ABB RobotStudio station: Lab1.rsstnx

Station Lab1 (saved by RobotStudio 25.5.11605.0)
Controller IRB140_6_81
  mechanical unit ROB_1: IRB140_6_81_C_03, 6 joints, base frame (0, 0, 0) mm
Layout (positions relative to the parent item):
  - IRB140_6_81_C_03 [mechanism, from %ABB.RobotStudio.Models.IRB140%\IRB140_6_81_C_G_03.rslib] at (0, 0, 0) mm; joint values [0, 0, 0, 0, 0.5236, 0] (rad or m)
  - MyNewTool [mechanism] at (506.29, 0, 679.5) mm, rotated rx 180 ry 60 rz 180 deg
      TCP MyNewTool at (110.98, -0.23, 41.34) mm, rotated rx 0 ry -30 rz 180 deg
      links: Assembly 2
  - Pastel [part] at (327.56, -460.42, -59) mm, rotated rx 180 ry 0 rz -90 deg, size 150 x 200 x 50 mm
  - Banda [smart component]
      signals: DI DI_01, DI DI_02
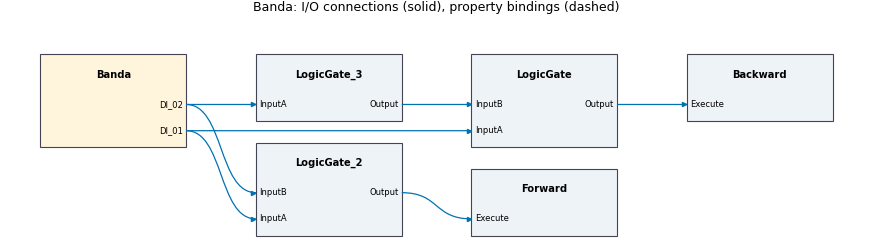
      connections:
        Banda.DI_02 -> LogicGate_3.InputA
        LogicGate_3.Output -> LogicGate.InputB
        LogicGate.Output -> Backward.Execute
        Banda.DI_02 -> LogicGate_2.InputB
        LogicGate_2.Output -> Forward.Execute
        Banda.DI_01 -> LogicGate_2.InputA
        Banda.DI_01 -> LogicGate.InputA
    - LogicGate [smart component, from Components\LogicGate.rslib]
        properties: Operator=AND; Delay=0.4
    - LogicGate_2 [smart component, from Components\LogicGate.rslib]
        properties: Operator=AND; Delay=0.4
    - LogicGate_3 [smart component, from Components\LogicGate.rslib]
        properties: Operator=NOT; Delay=0
    - Forward [smart component, from Components\LinearMover.rslib]
        properties: Object=Pastel; Direction=[0 -0.001 0]; Speed=0.328; Reference=Local; ReferenceObject=(none)
    - Backward [smart component, from Components\LinearMover.rslib]
        properties: Object=Pastel; Direction=[0 0.001 0]; Speed=0.328; Reference=Local; ReferenceObject=(none)
    - Start [smart component, from Components\Positioner.rslib] at (0, 0, 0) mm
        properties: Object=Pastel; Position=[-0.845372 -0.460416 -0.059]; Orientation=[3.14159265358979 0 -1.5707963267949]; Reference=Global; ReferenceObject=(none)
    - End [smart component, from Components\Positioner.rslib]
        properties: Object=Pastel; Position=[0.014628 -0.460416 -0.059]; Orientation=[3.14159265358979 0 -1.5707963267949]; Reference=Global; ReferenceObject=(none)
Attachment: MyNewTool is attached to IRB140_6_81_C_03 / Link6
Attachment: Start is attached to IRB140_6_81_C_03 / Link6
Station signals: DI DI_01, DI DI_02, DI DI_03
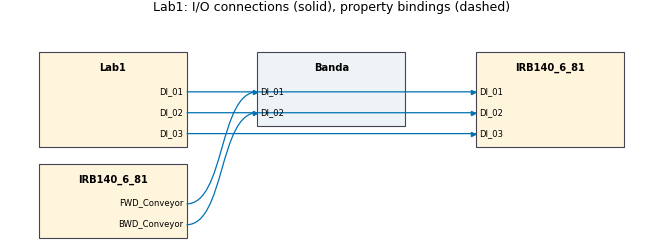
Station logic (signal -> signal, property => property):
  Lab1.DI_01 -> IRB140_6_81.DI_01
  Lab1.DI_02 -> IRB140_6_81.DI_02
  Lab1.DI_03 -> IRB140_6_81.DI_03
  IRB140_6_81.FWD_Conveyor -> Banda.DI_01
  IRB140_6_81.BWD_Conveyor -> Banda.DI_02
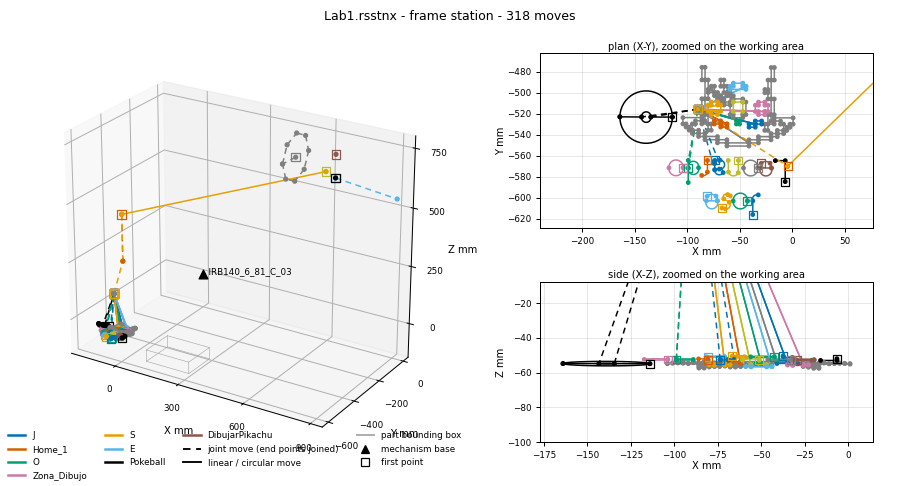
[picture p0: tool path of Lab1.rsstnx in frame station, 318 of 318 moves have a stored position in this frame; points joined in program order, loops and branches not executed]
Targets, tools, work objects and paths stored in the station, written as RAPID:
! task T_ROB1
MODULE Module1
  CONST robtarget E6_21:=[[119.525,55.911,0],[0,0,0,1],[0,0,0,0],[9E+09,9E+09,9E+09,9E+09,9E+09,9E+09]];
  PERS tooldata MyNewTool:=[TRUE,[[41.338,0.233,110.975],[0.866025404,0,0.5,0]],[1,[0,0,1],[1,0,0,0],0,0,0]];
  TASK PERS wobjdata Workobject_1:=[FALSE,TRUE,"",[[10.169850696,-448.889900169,-59],[0.018985691,0.705924683,-0.707820682,0.017313792]],[[0,0,0],[1,0,0,0]]];
  CONST robtarget D1:=[[123.545,108.722,0],[0,0,0,1],[-1,0,-1,1],[9E+09,9E+09,9E+09,9E+09,9E+09,9E+09]];
  CONST robtarget D2:=[[129.593,104.085,0],[0,0,0,1],[-1,0,-1,1],[9E+09,9E+09,9E+09,9E+09,9E+09,9E+09]];
  CONST robtarget D3:=[[123.185,98.948,0],[0,0,0,1],[-1,0,-1,1],[9E+09,9E+09,9E+09,9E+09,9E+09,9E+09]];
  CONST robtarget D4:=[[117.051,103.638,0],[0,0,0,1],[-1,0,-1,1],[9E+09,9E+09,9E+09,9E+09,9E+09,9E+09]];
  CONST robtarget Dibujo:=[[75,100,-150],[0,0,0,1],[-1,0,-1,1],[9E+09,9E+09,9E+09,9E+09,9E+09,9E+09]];
  CONST robtarget D5:=[[116.175,108.722,0],[0,0,0,1],[-1,0,-1,1],[9E+09,9E+09,9E+09,9E+09,9E+09,9E+09]];
  CONST robtarget D6:=[[137.325,108.722,0],[0,0,0,1],[-1,0,-1,1],[9E+09,9E+09,9E+09,9E+09,9E+09,9E+09]];
  CONST robtarget O1_2:=[[123.237,42.561,0],[0,0,0,1],[-1,0,-1,1],[9E+09,9E+09,9E+09,9E+09,9E+09,9E+09]];
  CONST robtarget O2_2:=[[130.813,49.503,0],[0,0,0,1],[-1,0,-1,1],[9E+09,9E+09,9E+09,9E+09,9E+09,9E+09]];
  CONST robtarget O3_2:=[[123.305,56.117,0],[0,0,0,1],[-1,0,-1,1],[9E+09,9E+09,9E+09,9E+09,9E+09,9E+09]];
  CONST robtarget O4_2:=[[115.831,49.349,0],[0,0,0,1],[-1,0,-1,1],[9E+09,9E+09,9E+09,9E+09,9E+09,9E+09]];
  CONST robtarget DibujoPk:=[[75,100,-150],[0,0,0,1],[0,0,0,0],[9E+09,9E+09,9E+09,9E+09,9E+09,9E+09]];
  CONST robtarget P2_1:=[[60.375,65.975,0],[0,0,0,1],[0,0,0,0],[9E+09,9E+09,9E+09,9E+09,9E+09,9E+09]];
  CONST robtarget P2_2:=[[60.375,56.975,0],[0,0,0,1],[0,0,0,0],[9E+09,9E+09,9E+09,9E+09,9E+09,9E+09]];
  CONST robtarget P2_3:=[[69.375,56.975,0],[0,0,0,1],[0,0,0,0],[9E+09,9E+09,9E+09,9E+09,9E+09,9E+09]];
  CONST robtarget P2_4:=[[69.375,65.975,0],[0,0,0,1],[0,0,0,0],[9E+09,9E+09,9E+09,9E+09,9E+09,9E+09]];
  CONST robtarget N1:=[[116.175,60.996,0],[0,0,0,1],[-1,0,-1,1],[9E+09,9E+09,9E+09,9E+09,9E+09,9E+09]];
  CONST robtarget N2:=[[127.893,61.049,0],[0,0,0,1],[-1,0,-1,1],[9E+09,9E+09,9E+09,9E+09,9E+09,9E+09]];
  CONST robtarget N3:=[[130.813,65.927,0],[0,0,0,1],[-1,0,-1,1],[9E+09,9E+09,9E+09,9E+09,9E+09,9E+09]];
  CONST robtarget N4:=[[127.169,70.439,0],[0,0,0,1],[-1,0,-1,1],[9E+09,9E+09,9E+09,9E+09,9E+09,9E+09]];
  CONST robtarget N5:=[[116.175,70.686,0],[0,0,0,1],[-1,0,-1,1],[9E+09,9E+09,9E+09,9E+09,9E+09,9E+09]];
  CONST robtarget P4_1:=[[81.375,71.975,0],[0,0,0,1],[0,0,0,0],[9E+09,9E+09,9E+09,9E+09,9E+09,9E+09]];
  CONST robtarget P4_2:=[[81.375,77.975,0],[0,0,0,1],[0,0,0,0],[9E+09,9E+09,9E+09,9E+09,9E+09,9E+09]];
  CONST robtarget P4_3:=[[78.375,77.975,0],[0,0,0,1],[0,0,0,0],[9E+09,9E+09,9E+09,9E+09,9E+09,9E+09]];
  CONST robtarget P4_4:=[[78.375,83.975,0],[0,0,0,1],[0,0,0,0],[9E+09,9E+09,9E+09,9E+09,9E+09,9E+09]];
  CONST robtarget P4_5:=[[81.375,83.975,0],[0,0,0,1],[0,0,0,0],[9E+09,9E+09,9E+09,9E+09,9E+09,9E+09]];
  CONST robtarget P4_6:=[[81.375,77.975,0],[0,0,0,1],[0,0,0,0],[9E+09,9E+09,9E+09,9E+09,9E+09,9E+09]];
  CONST robtarget P4_7:=[[84.375,77.975,0],[0,0,0,1],[0,0,0,0],[9E+09,9E+09,9E+09,9E+09,9E+09,9E+09]];
  CONST robtarget P4_8:=[[84.375,71.975,0],[0,0,0,1],[0,0,0,0],[9E+09,9E+09,9E+09,9E+09,9E+09,9E+09]];
  CONST robtarget P6_1:=[[69.375,35.975,0],[0,0,0,1],[0,0,0,0],[9E+09,9E+09,9E+09,9E+09,9E+09,9E+09]];
  CONST robtarget P6_2:=[[69.375,32.975,0],[0,0,0,1],[0,0,0,0],[9E+09,9E+09,9E+09,9E+09,9E+09,9E+09]];
  CONST robtarget P6_3:=[[63.375,32.975,0],[0,0,0,1],[0,0,0,0],[9E+09,9E+09,9E+09,9E+09,9E+09,9E+09]];
  CONST robtarget P6_4:=[[63.375,35.975,0],[0,0,0,1],[0,0,0,0],[9E+09,9E+09,9E+09,9E+09,9E+09,9E+09]];
  CONST robtarget P6_5:=[[60.375,35.975,0],[0,0,0,1],[0,0,0,0],[9E+09,9E+09,9E+09,9E+09,9E+09,9E+09]];
  CONST robtarget P6_6:=[[60.375,41.975,0],[0,0,0,1],[0,0,0,0],[9E+09,9E+09,9E+09,9E+09,9E+09,9E+09]];
  CONST robtarget P6_7:=[[63.375,41.975,0],[0,0,0,1],[0,0,0,0],[9E+09,9E+09,9E+09,9E+09,9E+09,9E+09]];
  CONST robtarget P6_8:=[[63.375,44.975,0],[0,0,0,1],[0,0,0,0],[9E+09,9E+09,9E+09,9E+09,9E+09,9E+09]];
  CONST robtarget P6_9:=[[69.375,44.975,0],[0,0,0,1],[0,0,0,0],[9E+09,9E+09,9E+09,9E+09,9E+09,9E+09]];
  CONST robtarget P6_10:=[[69.375,41.975,0],[0,0,0,1],[0,0,0,0],[9E+09,9E+09,9E+09,9E+09,9E+09,9E+09]];
  CONST robtarget P6_11:=[[72.375,41.975,0],[0,0,0,1],[0,0,0,0],[9E+09,9E+09,9E+09,9E+09,9E+09,9E+09]];
  CONST robtarget P6_12:=[[72.375,35.975,0],[0,0,0,1],[0,0,0,0],[9E+09,9E+09,9E+09,9E+09,9E+09,9E+09]];
  CONST robtarget O1_3:=[[123.237,113.603,0],[0,0,0,1],[-1,0,-1,1],[9E+09,9E+09,9E+09,9E+09,9E+09,9E+09]];
  CONST robtarget O2_3:=[[130.813,120.543,0],[0,0,0,1],[-1,0,-1,1],[9E+09,9E+09,9E+09,9E+09,9E+09,9E+09]];
  CONST robtarget O3_3:=[[123.305,127.159,0],[0,0,0,1],[-1,0,-1,1],[9E+09,9E+09,9E+09,9E+09,9E+09,9E+09]];
  CONST robtarget O4_3:=[[115.831,120.388,0],[0,0,0,1],[-1,0,-1,1],[9E+09,9E+09,9E+09,9E+09,9E+09,9E+09]];
  CONST robtarget PB1:=[[74.913,124.015,0],[0,0,0,1],[-1,0,-1,1],[9E+09,9E+09,9E+09,9E+09,9E+09,9E+09]];
  CONST robtarget PB2:=[[100,149.015,0],[0,0,0,1],[-1,0,-1,1],[9E+09,9E+09,9E+09,9E+09,9E+09,9E+09]];
  CONST robtarget PB3:=[[74.812,174.015,0],[0,0,0,1],[-1,0,-1,1],[9E+09,9E+09,9E+09,9E+09,9E+09,9E+09]];
  CONST robtarget PB4:=[[50,149.015,0],[0,0,0,1],[-1,0,-1,1],[9E+09,9E+09,9E+09,9E+09,9E+09,9E+09]];
  CONST robtarget PB5:=[[74.913,144.515,0],[0,0,0,1],[-1,0,-1,1],[9E+09,9E+09,9E+09,9E+09,9E+09,9E+09]];
  CONST robtarget PB6:=[[80,149.015,0],[0,0,0,1],[-1,0,-1,1],[9E+09,9E+09,9E+09,9E+09,9E+09,9E+09]];
  CONST robtarget PB7:=[[74.913,153.345,0],[0,0,0,1],[-1,0,-1,1],[9E+09,9E+09,9E+09,9E+09,9E+09,9E+09]];
  CONST robtarget PB8:=[[70,149.015,0],[0,0,0,1],[-1,0,-1,1],[9E+09,9E+09,9E+09,9E+09,9E+09,9E+09]];
  CONST robtarget J1:=[[167.685,47.174,0],[0,0,0,1],[-1,0,-1,1],[9E+09,9E+09,9E+09,9E+09,9E+09,9E+09]];
  CONST robtarget J2:=[[154.611,47.174,0],[0,0,0,1],[-1,0,-1,1],[9E+09,9E+09,9E+09,9E+09,9E+09,9E+09]];
  CONST robtarget J3:=[[150.083,46.324,0],[0,0,0,1],[-1,0,-1,1],[9E+09,9E+09,9E+09,9E+09,9E+09,9E+09]];
  CONST robtarget J4:=[[148.923,41.986,0],[0,0,0,1],[-1,0,-1,1],[9E+09,9E+09,9E+09,9E+09,9E+09,9E+09]];
  CONST robtarget P8_1:=[[45.375,53.975,0],[0,0,0,1],[0,0,0,0],[9E+09,9E+09,9E+09,9E+09,9E+09,9E+09]];
  CONST robtarget P8_2:=[[45.375,56.975,0],[0,0,0,1],[0,0,0,0],[9E+09,9E+09,9E+09,9E+09,9E+09,9E+09]];
  CONST robtarget P8_3:=[[42.375,56.975,0],[0,0,0,1],[0,0,0,0],[9E+09,9E+09,9E+09,9E+09,9E+09,9E+09]];
  CONST robtarget P8_4:=[[42.375,65.975,0],[0,0,0,1],[0,0,0,0],[9E+09,9E+09,9E+09,9E+09,9E+09,9E+09]];
  CONST robtarget P8_5:=[[45.375,65.975,0],[0,0,0,1],[0,0,0,0],[9E+09,9E+09,9E+09,9E+09,9E+09,9E+09]];
  CONST robtarget P8_6:=[[45.375,68.975,0],[0,0,0,1],[0,0,0,0],[9E+09,9E+09,9E+09,9E+09,9E+09,9E+09]];
  CONST robtarget P8_7:=[[48.375,68.975,0],[0,0,0,1],[0,0,0,0],[9E+09,9E+09,9E+09,9E+09,9E+09,9E+09]];
  CONST robtarget P8_8:=[[48.375,53.975,0],[0,0,0,1],[0,0,0,0],[9E+09,9E+09,9E+09,9E+09,9E+09,9E+09]];
  CONST robtarget wobjreal:=[[10.17,-448.89,43.77],[0.275144,0.645288,0.659942,-0.269026],[-1,0,0,1],[9E+09,9E+09,9E+09,9E+09,9E+09,9E+09]];
  CONST robtarget P1_1:=[[99.375,50.975,0],[0,0,0,1],[0,0,0,0],[9E+09,9E+09,9E+09,9E+09,9E+09,9E+09]];
  CONST robtarget P1_2:=[[99.375,41.975,0],[0,0,0,1],[0,0,0,0],[9E+09,9E+09,9E+09,9E+09,9E+09,9E+09]];
  CONST robtarget P1_3:=[[96.375,41.975,0],[0,0,0,1],[0,0,0,0],[9E+09,9E+09,9E+09,9E+09,9E+09,9E+09]];
  CONST robtarget P1_4:=[[96.375,29.975,0],[0,0,0,1],[0,0,0,0],[9E+09,9E+09,9E+09,9E+09,9E+09,9E+09]];
  CONST robtarget P1_5:=[[93.375,29.975,0],[0,0,0,1],[0,0,0,0],[9E+09,9E+09,9E+09,9E+09,9E+09,9E+09]];
  CONST robtarget P1_6:=[[93.375,23.975,0],[0,0,0,1],[0,0,0,0],[9E+09,9E+09,9E+09,9E+09,9E+09,9E+09]];
  CONST robtarget P1_7:=[[90.375,23.975,0],[0,0,0,1],[0,0,0,0],[9E+09,9E+09,9E+09,9E+09,9E+09,9E+09]];
  CONST robtarget P1_8:=[[90.375,17.975,0],[0,0,0,1],[0,0,0,0],[9E+09,9E+09,9E+09,9E+09,9E+09,9E+09]];
  CONST robtarget P1_9:=[[87.375,17.975,0],[0,0,0,1],[0,0,0,0],[9E+09,9E+09,9E+09,9E+09,9E+09,9E+09]];
  CONST robtarget P1_10:=[[87.375,14.975,0],[0,0,0,1],[0,0,0,0],[9E+09,9E+09,9E+09,9E+09,9E+09,9E+09]];
  CONST robtarget P1_11:=[[84.375,14.975,0],[0,0,0,1],[0,0,0,0],[9E+09,9E+09,9E+09,9E+09,9E+09,9E+09]];
  CONST robtarget P1_12:=[[84.375,11.975,0],[0,0,0,1],[0,0,0,0],[9E+09,9E+09,9E+09,9E+09,9E+09,9E+09]];
  CONST robtarget P1_13:=[[81.375,11.975,0],[0,0,0,1],[0,0,0,0],[9E+09,9E+09,9E+09,9E+09,9E+09,9E+09]];
  CONST robtarget P1_14:=[[81.375,8.975,0],[0,0,0,1],[0,0,0,0],[9E+09,9E+09,9E+09,9E+09,9E+09,9E+09]];
  CONST robtarget P1_15:=[[75.375,8.975,0],[0,0,0,1],[0,0,0,0],[9E+09,9E+09,9E+09,9E+09,9E+09,9E+09]];
  CONST robtarget P1_16:=[[75.375,26.975,0],[0,0,0,1],[0,0,0,0],[9E+09,9E+09,9E+09,9E+09,9E+09,9E+09]];
  CONST robtarget P1_17:=[[78.375,26.975,0],[0,0,0,1],[0,0,0,0],[9E+09,9E+09,9E+09,9E+09,9E+09,9E+09]];
  CONST robtarget P1_18:=[[78.375,29.975,0],[0,0,0,1],[0,0,0,0],[9E+09,9E+09,9E+09,9E+09,9E+09,9E+09]];
  CONST robtarget P1_19:=[[72.375,29.975,0],[0,0,0,1],[0,0,0,0],[9E+09,9E+09,9E+09,9E+09,9E+09,9E+09]];
  CONST robtarget P1_20:=[[72.375,26.975,0],[0,0,0,1],[0,0,0,0],[9E+09,9E+09,9E+09,9E+09,9E+09,9E+09]];
  CONST robtarget P1_21:=[[57.375,26.975,0],[0,0,0,1],[0,0,0,0],[9E+09,9E+09,9E+09,9E+09,9E+09,9E+09]];
  CONST robtarget P1_22:=[[57.375,29.975,0],[0,0,0,1],[0,0,0,0],[9E+09,9E+09,9E+09,9E+09,9E+09,9E+09]];
  CONST robtarget P1_23:=[[39.375,29.975,0],[0,0,0,1],[0,0,0,0],[9E+09,9E+09,9E+09,9E+09,9E+09,9E+09]];
  CONST robtarget P1_24:=[[39.375,26.975,0],[0,0,0,1],[0,0,0,0],[9E+09,9E+09,9E+09,9E+09,9E+09,9E+09]];
  CONST robtarget P1_25:=[[27.375,26.975,0],[0,0,0,1],[0,0,0,0],[9E+09,9E+09,9E+09,9E+09,9E+09,9E+09]];
  CONST robtarget P1_26:=[[27.375,29.975,0],[0,0,0,1],[0,0,0,0],[9E+09,9E+09,9E+09,9E+09,9E+09,9E+09]];
  CONST robtarget P1_27:=[[39.375,29.975,0],[0,0,0,1],[0,0,0,0],[9E+09,9E+09,9E+09,9E+09,9E+09,9E+09]];
  CONST robtarget P1_28:=[[39.375,32.975,0],[0,0,0,1],[0,0,0,0],[9E+09,9E+09,9E+09,9E+09,9E+09,9E+09]];
  CONST robtarget P1_29:=[[48.375,32.975,0],[0,0,0,1],[0,0,0,0],[9E+09,9E+09,9E+09,9E+09,9E+09,9E+09]];
  CONST robtarget P1_30:=[[48.375,35.975,0],[0,0,0,1],[0,0,0,0],[9E+09,9E+09,9E+09,9E+09,9E+09,9E+09]];
  CONST robtarget P1_31:=[[51.375,35.975,0],[0,0,0,1],[0,0,0,0],[9E+09,9E+09,9E+09,9E+09,9E+09,9E+09]];
  CONST robtarget P1_32:=[[51.375,32.975,0],[0,0,0,1],[0,0,0,0],[9E+09,9E+09,9E+09,9E+09,9E+09,9E+09]];
  CONST robtarget P1_33:=[[57.375,32.975,0],[0,0,0,1],[0,0,0,0],[9E+09,9E+09,9E+09,9E+09,9E+09,9E+09]];
  CONST robtarget P1_34:=[[57.375,29.975,0],[0,0,0,1],[0,0,0,0],[9E+09,9E+09,9E+09,9E+09,9E+09,9E+09]];
  CONST robtarget P1_35:=[[72.375,29.975,0],[0,0,0,1],[0,0,0,0],[9E+09,9E+09,9E+09,9E+09,9E+09,9E+09]];
  CONST robtarget P1_36:=[[72.375,32.975,0],[0,0,0,1],[0,0,0,0],[9E+09,9E+09,9E+09,9E+09,9E+09,9E+09]];
  CONST robtarget P1_37:=[[81.375,32.975,0],[0,0,0,1],[0,0,0,0],[9E+09,9E+09,9E+09,9E+09,9E+09,9E+09]];
  CONST robtarget P1_38:=[[81.375,35.975,0],[0,0,0,1],[0,0,0,0],[9E+09,9E+09,9E+09,9E+09,9E+09,9E+09]];
  CONST robtarget P1_39:=[[87.375,35.975,0],[0,0,0,1],[0,0,0,0],[9E+09,9E+09,9E+09,9E+09,9E+09,9E+09]];
  CONST robtarget P1_40:=[[87.375,32.975,0],[0,0,0,1],[0,0,0,0],[9E+09,9E+09,9E+09,9E+09,9E+09,9E+09]];
  CONST robtarget P1_41:=[[81.375,32.975,0],[0,0,0,1],[0,0,0,0],[9E+09,9E+09,9E+09,9E+09,9E+09,9E+09]];
  CONST robtarget P1_42:=[[81.375,26.975,0],[0,0,0,1],[0,0,0,0],[9E+09,9E+09,9E+09,9E+09,9E+09,9E+09]];
  CONST robtarget P1_43:=[[78.375,26.975,0],[0,0,0,1],[0,0,0,0],[9E+09,9E+09,9E+09,9E+09,9E+09,9E+09]];
  CONST robtarget P1_44:=[[78.375,20.975,0],[0,0,0,1],[0,0,0,0],[9E+09,9E+09,9E+09,9E+09,9E+09,9E+09]];
  CONST robtarget P1_45:=[[81.375,20.975,0],[0,0,0,1],[0,0,0,0],[9E+09,9E+09,9E+09,9E+09,9E+09,9E+09]];
  CONST robtarget P1_46:=[[81.375,17.975,0],[0,0,0,1],[0,0,0,0],[9E+09,9E+09,9E+09,9E+09,9E+09,9E+09]];
  CONST robtarget P1_47:=[[87.375,17.975,0],[0,0,0,1],[0,0,0,0],[9E+09,9E+09,9E+09,9E+09,9E+09,9E+09]];
  CONST robtarget P1_48:=[[87.375,23.975,0],[0,0,0,1],[0,0,0,0],[9E+09,9E+09,9E+09,9E+09,9E+09,9E+09]];
  CONST robtarget P1_49:=[[90.375,23.975,0],[0,0,0,1],[0,0,0,0],[9E+09,9E+09,9E+09,9E+09,9E+09,9E+09]];
  CONST robtarget P1_50:=[[90.375,29.975,0],[0,0,0,1],[0,0,0,0],[9E+09,9E+09,9E+09,9E+09,9E+09,9E+09]];
  CONST robtarget P1_51:=[[93.375,29.975,0],[0,0,0,1],[0,0,0,0],[9E+09,9E+09,9E+09,9E+09,9E+09,9E+09]];
  CONST robtarget P1_52:=[[93.375,41.975,0],[0,0,0,1],[0,0,0,0],[9E+09,9E+09,9E+09,9E+09,9E+09,9E+09]];
  CONST robtarget P1_53:=[[96.375,41.975,0],[0,0,0,1],[0,0,0,0],[9E+09,9E+09,9E+09,9E+09,9E+09,9E+09]];
  CONST robtarget P1_54:=[[96.375,50.975,0],[0,0,0,1],[0,0,0,0],[9E+09,9E+09,9E+09,9E+09,9E+09,9E+09]];
  CONST robtarget P1_55:=[[99.375,50.975,0],[0,0,0,1],[0,0,0,0],[9E+09,9E+09,9E+09,9E+09,9E+09,9E+09]];
  CONST robtarget P1_56:=[[99.375,71.975,0],[0,0,0,1],[0,0,0,0],[9E+09,9E+09,9E+09,9E+09,9E+09,9E+09]];
  CONST robtarget P1_57:=[[96.375,71.975,0],[0,0,0,1],[0,0,0,0],[9E+09,9E+09,9E+09,9E+09,9E+09,9E+09]];
  CONST robtarget P1_58:=[[96.375,80.975,0],[0,0,0,1],[0,0,0,0],[9E+09,9E+09,9E+09,9E+09,9E+09,9E+09]];
  CONST robtarget P1_59:=[[93.375,80.975,0],[0,0,0,1],[0,0,0,0],[9E+09,9E+09,9E+09,9E+09,9E+09,9E+09]];
  CONST robtarget P1_60:=[[93.375,92.975,0],[0,0,0,1],[0,0,0,0],[9E+09,9E+09,9E+09,9E+09,9E+09,9E+09]];
  CONST robtarget P1_61:=[[90.375,92.975,0],[0,0,0,1],[0,0,0,0],[9E+09,9E+09,9E+09,9E+09,9E+09,9E+09]];
  CONST robtarget P1_62:=[[90.375,98.975,0],[0,0,0,1],[0,0,0,0],[9E+09,9E+09,9E+09,9E+09,9E+09,9E+09]];
  CONST robtarget P1_63:=[[87.375,98.975,0],[0,0,0,1],[0,0,0,0],[9E+09,9E+09,9E+09,9E+09,9E+09,9E+09]];
  CONST robtarget P1_64:=[[87.375,104.975,0],[0,0,0,1],[0,0,0,0],[9E+09,9E+09,9E+09,9E+09,9E+09,9E+09]];
  CONST robtarget P1_65:=[[81.375,104.975,0],[0,0,0,1],[0,0,0,0],[9E+09,9E+09,9E+09,9E+09,9E+09,9E+09]];
  CONST robtarget P1_66:=[[81.375,101.975,0],[0,0,0,1],[0,0,0,0],[9E+09,9E+09,9E+09,9E+09,9E+09,9E+09]];
  CONST robtarget P1_67:=[[78.375,101.975,0],[0,0,0,1],[0,0,0,0],[9E+09,9E+09,9E+09,9E+09,9E+09,9E+09]];
  CONST robtarget P1_68:=[[78.375,95.975,0],[0,0,0,1],[0,0,0,0],[9E+09,9E+09,9E+09,9E+09,9E+09,9E+09]];
  CONST robtarget P1_69:=[[81.375,95.975,0],[0,0,0,1],[0,0,0,0],[9E+09,9E+09,9E+09,9E+09,9E+09,9E+09]];
  CONST robtarget P1_70:=[[81.375,89.975,0],[0,0,0,1],[0,0,0,0],[9E+09,9E+09,9E+09,9E+09,9E+09,9E+09]];
  CONST robtarget P1_71:=[[87.375,89.975,0],[0,0,0,1],[0,0,0,0],[9E+09,9E+09,9E+09,9E+09,9E+09,9E+09]];
  CONST robtarget P1_72:=[[87.375,86.975,0],[0,0,0,1],[0,0,0,0],[9E+09,9E+09,9E+09,9E+09,9E+09,9E+09]];
  CONST robtarget P1_73:=[[81.375,86.975,0],[0,0,0,1],[0,0,0,0],[9E+09,9E+09,9E+09,9E+09,9E+09,9E+09]];
  CONST robtarget P1_74:=[[81.375,89.975,0],[0,0,0,1],[0,0,0,0],[9E+09,9E+09,9E+09,9E+09,9E+09,9E+09]];
  CONST robtarget P1_75:=[[72.375,89.975,0],[0,0,0,1],[0,0,0,0],[9E+09,9E+09,9E+09,9E+09,9E+09,9E+09]];
  CONST robtarget P1_76:=[[72.375,92.975,0],[0,0,0,1],[0,0,0,0],[9E+09,9E+09,9E+09,9E+09,9E+09,9E+09]];
  CONST robtarget P1_77:=[[57.375,92.975,0],[0,0,0,1],[0,0,0,0],[9E+09,9E+09,9E+09,9E+09,9E+09,9E+09]];
  CONST robtarget P1_78:=[[57.375,89.975,0],[0,0,0,1],[0,0,0,0],[9E+09,9E+09,9E+09,9E+09,9E+09,9E+09]];
  CONST robtarget P1_79:=[[51.375,89.975,0],[0,0,0,1],[0,0,0,0],[9E+09,9E+09,9E+09,9E+09,9E+09,9E+09]];
  CONST robtarget P1_80:=[[51.375,83.975,0],[0,0,0,1],[0,0,0,0],[9E+09,9E+09,9E+09,9E+09,9E+09,9E+09]];
  CONST robtarget P1_81:=[[54.375,83.975,0],[0,0,0,1],[0,0,0,0],[9E+09,9E+09,9E+09,9E+09,9E+09,9E+09]];
  CONST robtarget P1_82:=[[54.375,80.975,0],[0,0,0,1],[0,0,0,0],[9E+09,9E+09,9E+09,9E+09,9E+09,9E+09]];
  CONST robtarget P1_83:=[[57.375,80.975,0],[0,0,0,1],[0,0,0,0],[9E+09,9E+09,9E+09,9E+09,9E+09,9E+09]];
  CONST robtarget P1_84:=[[57.375,77.975,0],[0,0,0,1],[0,0,0,0],[9E+09,9E+09,9E+09,9E+09,9E+09,9E+09]];
  CONST robtarget P1_85:=[[60.375,77.975,0],[0,0,0,1],[0,0,0,0],[9E+09,9E+09,9E+09,9E+09,9E+09,9E+09]];
  CONST robtarget P1_86:=[[60.375,74.975,0],[0,0,0,1],[0,0,0,0],[9E+09,9E+09,9E+09,9E+09,9E+09,9E+09]];
  CONST robtarget P1_87:=[[63.375,74.975,0],[0,0,0,1],[0,0,0,0],[9E+09,9E+09,9E+09,9E+09,9E+09,9E+09]];
  CONST robtarget P1_88:=[[63.375,68.975,0],[0,0,0,1],[0,0,0,0],[9E+09,9E+09,9E+09,9E+09,9E+09,9E+09]];
  CONST robtarget P1_89:=[[72.375,68.975,0],[0,0,0,1],[0,0,0,0],[9E+09,9E+09,9E+09,9E+09,9E+09,9E+09]];
  CONST robtarget P1_90:=[[72.375,65.975,0],[0,0,0,1],[0,0,0,0],[9E+09,9E+09,9E+09,9E+09,9E+09,9E+09]];
  CONST robtarget P1_91:=[[75.375,65.975,0],[0,0,0,1],[0,0,0,0],[9E+09,9E+09,9E+09,9E+09,9E+09,9E+09]];
  CONST robtarget P1_92:=[[75.375,56.975,0],[0,0,0,1],[0,0,0,0],[9E+09,9E+09,9E+09,9E+09,9E+09,9E+09]];
  CONST robtarget P1_93:=[[72.375,56.975,0],[0,0,0,1],[0,0,0,0],[9E+09,9E+09,9E+09,9E+09,9E+09,9E+09]];
  CONST robtarget P1_94:=[[72.375,53.975,0],[0,0,0,1],[0,0,0,0],[9E+09,9E+09,9E+09,9E+09,9E+09,9E+09]];
  CONST robtarget P1_95:=[[60.375,53.975,0],[0,0,0,1],[0,0,0,0],[9E+09,9E+09,9E+09,9E+09,9E+09,9E+09]];
  CONST robtarget P1_96:=[[60.375,56.975,0],[0,0,0,1],[0,0,0,0],[9E+09,9E+09,9E+09,9E+09,9E+09,9E+09]];
  CONST robtarget P1_97:=[[57.375,56.975,0],[0,0,0,1],[0,0,0,0],[9E+09,9E+09,9E+09,9E+09,9E+09,9E+09]];
  CONST robtarget P1_98:=[[57.375,65.975,0],[0,0,0,1],[0,0,0,0],[9E+09,9E+09,9E+09,9E+09,9E+09,9E+09]];
  CONST robtarget P1_99:=[[54.375,65.975,0],[0,0,0,1],[0,0,0,0],[9E+09,9E+09,9E+09,9E+09,9E+09,9E+09]];
  CONST robtarget P1_100:=[[54.375,68.975,0],[0,0,0,1],[0,0,0,0],[9E+09,9E+09,9E+09,9E+09,9E+09,9E+09]];
  CONST robtarget P1_101:=[[51.375,68.975,0],[0,0,0,1],[0,0,0,0],[9E+09,9E+09,9E+09,9E+09,9E+09,9E+09]];
  CONST robtarget P1_102:=[[51.375,71.975,0],[0,0,0,1],[0,0,0,0],[9E+09,9E+09,9E+09,9E+09,9E+09,9E+09]];
  CONST robtarget P1_103:=[[45.375,71.975,0],[0,0,0,1],[0,0,0,0],[9E+09,9E+09,9E+09,9E+09,9E+09,9E+09]];
  CONST robtarget P1_104:=[[45.375,74.975,0],[0,0,0,1],[0,0,0,0],[9E+09,9E+09,9E+09,9E+09,9E+09,9E+09]];
  CONST robtarget P1_105:=[[39.375,74.975,0],[0,0,0,1],[0,0,0,0],[9E+09,9E+09,9E+09,9E+09,9E+09,9E+09]];
  CONST robtarget P1_106:=[[39.375,77.975,0],[0,0,0,1],[0,0,0,0],[9E+09,9E+09,9E+09,9E+09,9E+09,9E+09]];
  CONST robtarget P1_107:=[[45.375,77.975,0],[0,0,0,1],[0,0,0,0],[9E+09,9E+09,9E+09,9E+09,9E+09,9E+09]];
  CONST robtarget P1_108:=[[45.375,74.975,0],[0,0,0,1],[0,0,0,0],[9E+09,9E+09,9E+09,9E+09,9E+09,9E+09]];
  CONST robtarget P1_109:=[[51.375,74.975,0],[0,0,0,1],[0,0,0,0],[9E+09,9E+09,9E+09,9E+09,9E+09,9E+09]];
  CONST robtarget P1_110:=[[51.375,71.975,0],[0,0,0,1],[0,0,0,0],[9E+09,9E+09,9E+09,9E+09,9E+09,9E+09]];
  CONST robtarget P1_111:=[[54.375,71.975,0],[0,0,0,1],[0,0,0,0],[9E+09,9E+09,9E+09,9E+09,9E+09,9E+09]];
  CONST robtarget P1_112:=[[54.375,68.975,0],[0,0,0,1],[0,0,0,0],[9E+09,9E+09,9E+09,9E+09,9E+09,9E+09]];
  CONST robtarget P1_113:=[[60.375,68.975,0],[0,0,0,1],[0,0,0,0],[9E+09,9E+09,9E+09,9E+09,9E+09,9E+09]];
  CONST robtarget P1_114:=[[60.375,74.975,0],[0,0,0,1],[0,0,0,0],[9E+09,9E+09,9E+09,9E+09,9E+09,9E+09]];
  CONST robtarget P1_115:=[[57.375,74.975,0],[0,0,0,1],[0,0,0,0],[9E+09,9E+09,9E+09,9E+09,9E+09,9E+09]];
  CONST robtarget P1_116:=[[57.375,77.975,0],[0,0,0,1],[0,0,0,0],[9E+09,9E+09,9E+09,9E+09,9E+09,9E+09]];
  CONST robtarget P1_117:=[[54.375,77.975,0],[0,0,0,1],[0,0,0,0],[9E+09,9E+09,9E+09,9E+09,9E+09,9E+09]];
  CONST robtarget P1_118:=[[54.375,80.975,0],[0,0,0,1],[0,0,0,0],[9E+09,9E+09,9E+09,9E+09,9E+09,9E+09]];
  CONST robtarget P1_119:=[[51.375,80.975,0],[0,0,0,1],[0,0,0,0],[9E+09,9E+09,9E+09,9E+09,9E+09,9E+09]];
  CONST robtarget P1_120:=[[51.375,83.975,0],[0,0,0,1],[0,0,0,0],[9E+09,9E+09,9E+09,9E+09,9E+09,9E+09]];
  CONST robtarget P1_121:=[[45.375,83.975,0],[0,0,0,1],[0,0,0,0],[9E+09,9E+09,9E+09,9E+09,9E+09,9E+09]];
  CONST robtarget P1_122:=[[45.375,86.975,0],[0,0,0,1],[0,0,0,0],[9E+09,9E+09,9E+09,9E+09,9E+09,9E+09]];
  CONST robtarget P1_123:=[[48.375,86.975,0],[0,0,0,1],[0,0,0,0],[9E+09,9E+09,9E+09,9E+09,9E+09,9E+09]];
  CONST robtarget P1_124:=[[48.375,89.975,0],[0,0,0,1],[0,0,0,0],[9E+09,9E+09,9E+09,9E+09,9E+09,9E+09]];
  CONST robtarget P1_125:=[[39.375,89.975,0],[0,0,0,1],[0,0,0,0],[9E+09,9E+09,9E+09,9E+09,9E+09,9E+09]];
  CONST robtarget P1_126:=[[39.375,92.975,0],[0,0,0,1],[0,0,0,0],[9E+09,9E+09,9E+09,9E+09,9E+09,9E+09]];
  CONST robtarget P1_127:=[[27.375,92.975,0],[0,0,0,1],[0,0,0,0],[9E+09,9E+09,9E+09,9E+09,9E+09,9E+09]];
  CONST robtarget P1_128:=[[27.375,95.975,0],[0,0,0,1],[0,0,0,0],[9E+09,9E+09,9E+09,9E+09,9E+09,9E+09]];
  CONST robtarget P1_129:=[[39.375,95.975,0],[0,0,0,1],[0,0,0,0],[9E+09,9E+09,9E+09,9E+09,9E+09,9E+09]];
  CONST robtarget P1_130:=[[39.375,92.975,0],[0,0,0,1],[0,0,0,0],[9E+09,9E+09,9E+09,9E+09,9E+09,9E+09]];
  CONST robtarget P1_131:=[[57.375,92.975,0],[0,0,0,1],[0,0,0,0],[9E+09,9E+09,9E+09,9E+09,9E+09,9E+09]];
  CONST robtarget P1_132:=[[57.375,95.975,0],[0,0,0,1],[0,0,0,0],[9E+09,9E+09,9E+09,9E+09,9E+09,9E+09]];
  CONST robtarget P1_133:=[[72.375,95.975,0],[0,0,0,1],[0,0,0,0],[9E+09,9E+09,9E+09,9E+09,9E+09,9E+09]];
  CONST robtarget P1_134:=[[72.375,92.975,0],[0,0,0,1],[0,0,0,0],[9E+09,9E+09,9E+09,9E+09,9E+09,9E+09]];
  CONST robtarget P1_135:=[[78.375,92.975,0],[0,0,0,1],[0,0,0,0],[9E+09,9E+09,9E+09,9E+09,9E+09,9E+09]];
  CONST robtarget P1_136:=[[78.375,95.975,0],[0,0,0,1],[0,0,0,0],[9E+09,9E+09,9E+09,9E+09,9E+09,9E+09]];
  CONST robtarget P1_137:=[[75.375,95.975,0],[0,0,0,1],[0,0,0,0],[9E+09,9E+09,9E+09,9E+09,9E+09,9E+09]];
  CONST robtarget P1_138:=[[75.375,113.975,0],[0,0,0,1],[0,0,0,0],[9E+09,9E+09,9E+09,9E+09,9E+09,9E+09]];
  CONST robtarget P1_139:=[[81.375,113.975,0],[0,0,0,1],[0,0,0,0],[9E+09,9E+09,9E+09,9E+09,9E+09,9E+09]];
  CONST robtarget P1_140:=[[81.375,110.975,0],[0,0,0,1],[0,0,0,0],[9E+09,9E+09,9E+09,9E+09,9E+09,9E+09]];
  CONST robtarget P1_141:=[[84.375,110.975,0],[0,0,0,1],[0,0,0,0],[9E+09,9E+09,9E+09,9E+09,9E+09,9E+09]];
  CONST robtarget P1_142:=[[84.375,107.975,0],[0,0,0,1],[0,0,0,0],[9E+09,9E+09,9E+09,9E+09,9E+09,9E+09]];
  CONST robtarget P1_143:=[[87.375,107.975,0],[0,0,0,1],[0,0,0,0],[9E+09,9E+09,9E+09,9E+09,9E+09,9E+09]];
  CONST robtarget P1_144:=[[87.375,104.975,0],[0,0,0,1],[0,0,0,0],[9E+09,9E+09,9E+09,9E+09,9E+09,9E+09]];
  CONST robtarget P1_145:=[[90.375,104.975,0],[0,0,0,1],[0,0,0,0],[9E+09,9E+09,9E+09,9E+09,9E+09,9E+09]];
  CONST robtarget P1_146:=[[90.375,98.975,0],[0,0,0,1],[0,0,0,0],[9E+09,9E+09,9E+09,9E+09,9E+09,9E+09]];
  CONST robtarget P1_147:=[[93.375,98.975,0],[0,0,0,1],[0,0,0,0],[9E+09,9E+09,9E+09,9E+09,9E+09,9E+09]];
  CONST robtarget P1_148:=[[93.375,92.975,0],[0,0,0,1],[0,0,0,0],[9E+09,9E+09,9E+09,9E+09,9E+09,9E+09]];
  CONST robtarget P1_149:=[[96.375,92.975,0],[0,0,0,1],[0,0,0,0],[9E+09,9E+09,9E+09,9E+09,9E+09,9E+09]];
  CONST robtarget P1_150:=[[96.375,80.975,0],[0,0,0,1],[0,0,0,0],[9E+09,9E+09,9E+09,9E+09,9E+09,9E+09]];
  CONST robtarget P1_151:=[[99.375,80.975,0],[0,0,0,1],[0,0,0,0],[9E+09,9E+09,9E+09,9E+09,9E+09,9E+09]];
  CONST robtarget P1_152:=[[99.375,71.975,0],[0,0,0,1],[0,0,0,0],[9E+09,9E+09,9E+09,9E+09,9E+09,9E+09]];
  CONST robtarget P1_153:=[[102.375,71.975,0],[0,0,0,1],[0,0,0,0],[9E+09,9E+09,9E+09,9E+09,9E+09,9E+09]];
  CONST robtarget P1_154:=[[102.375,50.975,0],[0,0,0,1],[0,0,0,0],[9E+09,9E+09,9E+09,9E+09,9E+09,9E+09]];
  CONST robtarget A1:=[[116.175,83.52,0],[0,0,0,1],[-1,0,-1,1],[9E+09,9E+09,9E+09,9E+09,9E+09,9E+09]];
  CONST robtarget A2:=[[125.057,83.52,0],[0,0,0,1],[-1,0,-1,1],[9E+09,9E+09,9E+09,9E+09,9E+09,9E+09]];
  CONST robtarget A3:=[[129.549,80.727,0],[0,0,0,1],[-1,0,-1,1],[9E+09,9E+09,9E+09,9E+09,9E+09,9E+09]];
  CONST robtarget A4:=[[127.721,75.478,0],[0,0,0,1],[-1,0,-1,1],[9E+09,9E+09,9E+09,9E+09,9E+09,9E+09]];
  CONST robtarget A5:=[[124.405,79.121,0],[0,0,0,1],[-1,0,-1,1],[9E+09,9E+09,9E+09,9E+09,9E+09,9E+09]];
  CONST robtarget A6:=[[119.869,74.173,0],[0,0,0,1],[-1,0,-1,1],[9E+09,9E+09,9E+09,9E+09,9E+09,9E+09]];
  CONST robtarget A7:=[[115.831,78.607,0],[0,0,0,1],[-1,0,-1,1],[9E+09,9E+09,9E+09,9E+09,9E+09,9E+09]];
  CONST robtarget A8:=[[116.673,81.448,0],[0,0,0,1],[-1,0,-1,1],[9E+09,9E+09,9E+09,9E+09,9E+09,9E+09]];
  CONST robtarget A9:=[[119.011,83.469,0],[0,0,0,1],[-1,0,-1,1],[9E+09,9E+09,9E+09,9E+09,9E+09,9E+09]];
  CONST robtarget L1:=[[136.191,16.345,0],[0,0,0,1],[-1,0,-1,1],[9E+09,9E+09,9E+09,9E+09,9E+09,9E+09]];
  CONST robtarget L2:=[[116.175,16.345,0],[0,0,0,1],[-1,0,-1,1],[9E+09,9E+09,9E+09,9E+09,9E+09,9E+09]];
  CONST robtarget L3:=[[116.175,25.793,0],[0,0,0,1],[-1,0,-1,1],[9E+09,9E+09,9E+09,9E+09,9E+09,9E+09]];
  CONST robtarget R1:=[[116.175,90.46,0],[0,0,0,1],[-1,0,-1,1],[9E+09,9E+09,9E+09,9E+09,9E+09,9E+09]];
  CONST robtarget R2:=[[127.309,90.513,0],[0,0,0,1],[-1,0,-1,1],[9E+09,9E+09,9E+09,9E+09,9E+09,9E+09]];
  CONST robtarget R2_2:=[[130.135,92.453,0],[0,0,0,1],[-1,-2,-2,0],[9E+09,9E+09,9E+09,9E+09,9E+09,9E+09]];
  CONST robtarget R3:=[[130.487,95.924,0],[0,0,0,1],[-1,0,-1,1],[9E+09,9E+09,9E+09,9E+09,9E+09,9E+09]];
  CONST robtarget P3_1:=[[81.375,44.975,0],[0,0,0,1],[0,0,0,0],[9E+09,9E+09,9E+09,9E+09,9E+09,9E+09]];
  CONST robtarget P3_2:=[[81.375,38.975,0],[0,0,0,1],[0,0,0,0],[9E+09,9E+09,9E+09,9E+09,9E+09,9E+09]];
  CONST robtarget P3_3:=[[78.375,38.975,0],[0,0,0,1],[0,0,0,0],[9E+09,9E+09,9E+09,9E+09,9E+09,9E+09]];
  CONST robtarget P3_4:=[[78.375,44.975,0],[0,0,0,1],[0,0,0,0],[9E+09,9E+09,9E+09,9E+09,9E+09,9E+09]];
  CONST robtarget P3_5:=[[81.375,44.975,0],[0,0,0,1],[0,0,0,0],[9E+09,9E+09,9E+09,9E+09,9E+09,9E+09]];
  CONST robtarget P3_6:=[[81.375,50.975,0],[0,0,0,1],[0,0,0,0],[9E+09,9E+09,9E+09,9E+09,9E+09,9E+09]];
  CONST robtarget P3_7:=[[84.375,50.975,0],[0,0,0,1],[0,0,0,0],[9E+09,9E+09,9E+09,9E+09,9E+09,9E+09]];
  CONST robtarget P3_8:=[[84.375,44.975,0],[0,0,0,1],[0,0,0,0],[9E+09,9E+09,9E+09,9E+09,9E+09,9E+09]];
  CONST robtarget S1:=[[161.551,76.518,0],[0,0,0,1],[-1,0,-1,1],[9E+09,9E+09,9E+09,9E+09,9E+09,9E+09]];
  CONST robtarget S2:=[[162.307,73.374,0],[0,0,0,1],[-1,0,-1,1],[9E+09,9E+09,9E+09,9E+09,9E+09,9E+09]];
  CONST robtarget S3:=[[159.977,69.026,0],[0,0,0,1],[-1,0,-1,1],[9E+09,9E+09,9E+09,9E+09,9E+09,9E+09]];
  CONST robtarget S4:=[[156.043,69.546,0],[0,0,0,1],[-1,0,-1,1],[9E+09,9E+09,9E+09,9E+09,9E+09,9E+09]];
  CONST robtarget S5:=[[152.747,74.93,0],[0,0,0,1],[-1,0,-1,1],[9E+09,9E+09,9E+09,9E+09,9E+09,9E+09]];
  CONST robtarget S6:=[[149.263,74.776,0],[0,0,0,1],[-1,0,-1,1],[9E+09,9E+09,9E+09,9E+09,9E+09,9E+09]];
  CONST robtarget S7:=[[148.697,71.136,0],[0,0,0,1],[-1,0,-1,1],[9E+09,9E+09,9E+09,9E+09,9E+09,9E+09]];
  CONST robtarget S8:=[[149.903,68.65,0],[0,0,0,1],[-1,0,-1,1],[9E+09,9E+09,9E+09,9E+09,9E+09,9E+09]];
  CONST robtarget Home_2:=[[138.534211034,14.836428397,-331.193016671],[0.001338278,-0.025663879,-0.001186167,0.999669029],[-2,0,-1,1],[9E+09,9E+09,9E+09,9E+09,9E+09,9E+09]];
  CONST robtarget Home:=[[148.797,15.297,-530.929],[0.001338278,-0.025663879,-0.001186167,0.999669029],[-1,-1,0,0],[9E+09,9E+09,9E+09,9E+09,9E+09,9E+09]];
  CONST robtarget O1:=[[154.731,52.294,0],[0,0,0,1],[-1,0,-1,1],[9E+09,9E+09,9E+09,9E+09,9E+09,9E+09]];
  CONST robtarget O2:=[[162.307,59.236,0],[0,0,0,1],[-1,0,-1,1],[9E+09,9E+09,9E+09,9E+09,9E+09,9E+09]];
  CONST robtarget O3:=[[154.799,65.85,0],[0,0,0,1],[-1,0,-1,1],[9E+09,9E+09,9E+09,9E+09,9E+09,9E+09]];
  CONST robtarget O4:=[[147.325,59.08,0],[0,0,0,1],[-1,0,-1,1],[9E+09,9E+09,9E+09,9E+09,9E+09,9E+09]];
  CONST robtarget P5_1:=[[78.375,59.975,0],[0,0,0,1],[0,0,0,0],[9E+09,9E+09,9E+09,9E+09,9E+09,9E+09]];
  CONST robtarget P5_2:=[[78.375,62.975,0],[0,0,0,1],[0,0,0,0],[9E+09,9E+09,9E+09,9E+09,9E+09,9E+09]];
  CONST robtarget P5_3:=[[81.375,62.975,0],[0,0,0,1],[0,0,0,0],[9E+09,9E+09,9E+09,9E+09,9E+09,9E+09]];
  CONST robtarget P5_4:=[[81.375,59.975,0],[0,0,0,1],[0,0,0,0],[9E+09,9E+09,9E+09,9E+09,9E+09,9E+09]];
  CONST robtarget Aura0:=[[-325.233,-481.73,-738.213],[0.707106781,0,0,0.707106781],[-1,-2,1,1],[9E+09,9E+09,9E+09,9E+09,9E+09,9E+09]];
  CONST robtarget Aura1:=[[-225.233,-481.73,-738.213],[0.707106781,0,0,0.707106781],[-1,-2,1,1],[9E+09,9E+09,9E+09,9E+09,9E+09,9E+09]];
  CONST robtarget Aura2:=[[-254.523,-481.73,-808.923],[0.707106781,0,0,0.707106781],[-1,0,3,0],[9E+09,9E+09,9E+09,9E+09,9E+09,9E+09]];
  CONST robtarget Aura3:=[[-325.233,-481.73,-838.213],[0.707106781,0,0,0.707106781],[-1,-2,1,1],[9E+09,9E+09,9E+09,9E+09,9E+09,9E+09]];
  CONST robtarget Aura4:=[[-395.943,-481.73,-808.923],[0.707106781,0,0,0.707106781],[0,-1,0,0],[9E+09,9E+09,9E+09,9E+09,9E+09,9E+09]];
  CONST robtarget Aura5:=[[-425.233,-481.73,-738.213],[0.707106781,0,0,0.707106781],[0,1,-2,1],[9E+09,9E+09,9E+09,9E+09,9E+09,9E+09]];
  CONST robtarget Aura6:=[[-395.943,-481.73,-667.503],[0.707106781,0,0,0.707106781],[0,-1,0,0],[9E+09,9E+09,9E+09,9E+09,9E+09,9E+09]];
  CONST robtarget Aura7:=[[-325.233,-481.73,-638.213],[0.707106781,0,0,0.707106781],[-1,-2,1,1],[9E+09,9E+09,9E+09,9E+09,9E+09,9E+09]];
  CONST robtarget Aura8:=[[-254.523,-481.73,-667.503],[0.707106781,0,0,0.707106781],[-1,0,-1,0],[9E+09,9E+09,9E+09,9E+09,9E+09,9E+09]];
  CONST robtarget P7_1:=[[69.375,80.975,0],[0,0,0,1],[0,0,0,0],[9E+09,9E+09,9E+09,9E+09,9E+09,9E+09]];
  CONST robtarget P7_2:=[[69.375,77.975,0],[0,0,0,1],[0,0,0,0],[9E+09,9E+09,9E+09,9E+09,9E+09,9E+09]];
  CONST robtarget P7_3:=[[63.375,77.975,0],[0,0,0,1],[0,0,0,0],[9E+09,9E+09,9E+09,9E+09,9E+09,9E+09]];
  CONST robtarget P7_4:=[[63.375,80.975,0],[0,0,0,1],[0,0,0,0],[9E+09,9E+09,9E+09,9E+09,9E+09,9E+09]];
  CONST robtarget P7_5:=[[60.375,80.975,0],[0,0,0,1],[0,0,0,0],[9E+09,9E+09,9E+09,9E+09,9E+09,9E+09]];
  CONST robtarget P7_6:=[[60.375,86.975,0],[0,0,0,1],[0,0,0,0],[9E+09,9E+09,9E+09,9E+09,9E+09,9E+09]];
  CONST robtarget P7_7:=[[63.375,86.975,0],[0,0,0,1],[0,0,0,0],[9E+09,9E+09,9E+09,9E+09,9E+09,9E+09]];
  CONST robtarget P7_8:=[[63.375,89.975,0],[0,0,0,1],[0,0,0,0],[9E+09,9E+09,9E+09,9E+09,9E+09,9E+09]];
  CONST robtarget P7_9:=[[69.375,89.975,0],[0,0,0,1],[0,0,0,0],[9E+09,9E+09,9E+09,9E+09,9E+09,9E+09]];
  CONST robtarget P7_10:=[[69.375,86.975,0],[0,0,0,1],[0,0,0,0],[9E+09,9E+09,9E+09,9E+09,9E+09,9E+09]];
  CONST robtarget P7_11:=[[72.375,86.975,0],[0,0,0,1],[0,0,0,0],[9E+09,9E+09,9E+09,9E+09,9E+09,9E+09]];
  CONST robtarget P7_12:=[[72.375,80.975,0],[0,0,0,1],[0,0,0,0],[9E+09,9E+09,9E+09,9E+09,9E+09,9E+09]];
  CONST robtarget E1:=[[150.297,90.658,0],[0,0,0,1],[-1,0,-1,1],[9E+09,9E+09,9E+09,9E+09,9E+09,9E+09]];
  CONST robtarget E2:=[[148.545,85.968,0],[0,0,0,1],[-1,0,-1,1],[9E+09,9E+09,9E+09,9E+09,9E+09,9E+09]];
  CONST robtarget E3:=[[150.177,82.248,0],[0,0,0,1],[-1,0,-1,1],[9E+09,9E+09,9E+09,9E+09,9E+09,9E+09]];
  CONST robtarget E4:=[[152.125,81.238,0],[0,0,0,1],[-1,0,-1,1],[9E+09,9E+09,9E+09,9E+09,9E+09,9E+09]];
  CONST robtarget E5:=[[154.713,80.9,0],[0,0,0,1],[-1,0,-1,1],[9E+09,9E+09,9E+09,9E+09,9E+09,9E+09]];
  CONST robtarget E6:=[[154.713,91.466,0],[0,0,0,1],[-1,0,-1,1],[9E+09,9E+09,9E+09,9E+09,9E+09,9E+09]];
  CONST robtarget E7:=[[162.307,85.934,0],[0,0,0,1],[-1,0,-1,1],[9E+09,9E+09,9E+09,9E+09,9E+09,9E+09]];
  CONST robtarget E1_2:=[[118.805,39.263,0],[0,0,0,1],[-1,0,-1,1],[9E+09,9E+09,9E+09,9E+09,9E+09,9E+09]];
  CONST robtarget E2_2:=[[117.051,34.573,0],[0,0,0,1],[-1,0,-1,1],[9E+09,9E+09,9E+09,9E+09,9E+09,9E+09]];
  CONST robtarget E3_2:=[[118.683,30.853,0],[0,0,0,1],[-1,0,-1,1],[9E+09,9E+09,9E+09,9E+09,9E+09,9E+09]];
  CONST robtarget E4_2:=[[120.645,29.839,0],[0,0,0,1],[-1,0,-1,1],[9E+09,9E+09,9E+09,9E+09,9E+09,9E+09]];
  CONST robtarget E5_2:=[[123.219,29.505,0],[0,0,0,1],[-1,0,-1,1],[9E+09,9E+09,9E+09,9E+09,9E+09,9E+09]];
  CONST robtarget E6_2:=[[123.219,40.071,0],[0,0,0,1],[-1,0,-1,1],[9E+09,9E+09,9E+09,9E+09,9E+09,9E+09]];
  CONST robtarget E7_2:=[[130.813,34.539,0],[0,0,0,1],[-1,-2,-2,0],[9E+09,9E+09,9E+09,9E+09,9E+09,9E+09]];
  CONST robtarget Home_F2:=[[-417.824726867,-613.120156159,-653.373090922],[0.678788419,0.165982914,-0.201536242,0.686352022],[-1,-1,0,1],[9E+09,9E+09,9E+09,9E+09,9E+09,9E+09]];
  CONST robtarget Mantenimiento:=[[-420.017689886,-888.965003638,-625.487828896],[0.678788419,0.165982914,-0.201536242,0.686352022],[0,0,0,0],[9E+09,9E+09,9E+09,9E+09,9E+09,9E+09]];
  CONST robtarget Home0:=[[-412.691499067,-612.89567271,-753.243004357],[0.678788419,0.165982914,-0.201536242,0.686352022],[-1,0,-1,0],[9E+09,9E+09,9E+09,9E+09,9E+09,9E+09]];
  CONST robtarget RealH:=[[-416.810979787,-568.840149732,-670.795454874],[0.707820682,-0.017313792,-0.018985691,0.705924683],[0,-1,0,0],[9E+09,9E+09,9E+09,9E+09,9E+09,9E+09]];
  PROC J()
    MoveJ J1,v100,z1,MyNewTool\WObj:=Workobject_1;
    MoveL J2,v100,z1,MyNewTool\WObj:=Workobject_1;
    MoveC J3,J4,v100,z1,MyNewTool\WObj:=Workobject_1;
  ENDPROC
  PROC Home_1()
    MoveJ Home,v100,z1,MyNewTool\WObj:=Workobject_1;
    MoveJ Home_2,v100,z1,MyNewTool\WObj:=Workobject_1;
  ENDPROC
  PROC main()
    Reset FWD_Conveyor;
    Reset BWD_Conveyor;
    Reset DO_01;
    Reset DO_02;
    Reset DO_03;
    Set BWD_Conveyor;
    Set FWD_Conveyor;
    WaitTime 2.591;
    Reset FWD_Conveyor;
    Reset BWD_Conveyor;
    Set DO_01;
    Real_Home;
    Home_1;
    Zona_Dibujo;
    J;
    Zona_Dibujo;
    O;
    Zona_Dibujo;
    S;
    Zona_Dibujo;
    E;
    Zona_Dibujo;
    L;
    Zona_Dibujo;
    E_2;
    Zona_Dibujo;
    O_2;
    Zona_Dibujo;
    N;
    Zona_Dibujo;
    A;
    Zona_Dibujo;
    R;
    Zona_Dibujo;
    D;
    Zona_Dibujo;
    O_3;
    Zona_Dibujo;
    Pokeball;
    Zona_Dibujo;
    DibujarPikachu;
    Reset DO_01;
    Home_F;
    Set BWD_Conveyor;
    Set FWD_Conveyor;
    WaitTime 1;
    Reset FWD_Conveyor;
    Reset BWD_Conveyor;
    Set DO_03;
    Real_Home;
    Aura;
    Real_Home;
    Reset DO_03;
    Set DO_02;
    Mantenimiento_p;
    Real_Home;
    Reset DO_02;
  ENDPROC
  PROC O()
    MoveJ O1,v100,z1,MyNewTool\WObj:=Workobject_1;
    MoveC O2,O3,v100,z1,MyNewTool\WObj:=Workobject_1;
    MoveC O4,O1,v100,z1,MyNewTool\WObj:=Workobject_1;
  ENDPROC
  PROC Zona_Dibujo()
    MoveJ Dibujo,v100,z1,MyNewTool\WObj:=Workobject_1;
  ENDPROC
  PROC S()
    MoveJ S1,v100,z1,MyNewTool\WObj:=Workobject_1;
    MoveL S2,v100,z1,MyNewTool\WObj:=Workobject_1;
    MoveC S3,S4,v100,z1,MyNewTool\WObj:=Workobject_1;
    MoveL S5,v100,z1,MyNewTool\WObj:=Workobject_1;
    MoveC S6,S7,v100,z1,MyNewTool\WObj:=Workobject_1;
    MoveL S8,v100,z1,MyNewTool\WObj:=Workobject_1;
  ENDPROC
  PROC E()
    MoveJ E1,v100,z1,MyNewTool\WObj:=Workobject_1;
    MoveC E2,E3,v100,z1,MyNewTool\WObj:=Workobject_1;
    MoveC E4,E5,v100,z1,MyNewTool\WObj:=Workobject_1;
    MoveL E6,v100,z1,MyNewTool\WObj:=Workobject_1;
    MoveC E7,E5,v100,z1,MyNewTool\WObj:=Workobject_1;
  ENDPROC
  PROC Pokeball()
    MoveJ PB1,v100,z1,MyNewTool\WObj:=Workobject_1;
    MoveC PB2,PB3,v100,z1,MyNewTool\WObj:=Workobject_1;
    MoveC PB4,PB1,v100,z1,MyNewTool\WObj:=Workobject_1;
    MoveL PB5,v100,z1,MyNewTool\WObj:=Workobject_1;
    MoveC PB6,PB7,v100,z1,MyNewTool\WObj:=Workobject_1;
    MoveC PB8,PB5,v100,z1,MyNewTool\WObj:=Workobject_1;
    MoveJ Dibujo,v100,z1,MyNewTool\WObj:=Workobject_1;
    MoveJ PB7,v100,z1,MyNewTool\WObj:=Workobject_1;
    MoveL PB3,v100,z1,MyNewTool\WObj:=Workobject_1;
  ENDPROC
  PROC DibujarPikachu()
    ConfJ \Off;
    ConfL \Off;
    Trazo1;
    Trazo2;
    Trazo3;
    Trazo4;
    Trazo5;
    Trazo6;
    Trazo7;
    Trazo8;
    MoveL DibujoPk,v100,z1,MyNewTool\WObj:=Workobject_1;
  ENDPROC
  PROC Trazo1()
    MoveL DibujoPk,v100,z1,MyNewTool\WObj:=Workobject_1;
    MoveL P1_1,v100,z1,MyNewTool\WObj:=Workobject_1;
    MoveL P1_2,v100,z1,MyNewTool\WObj:=Workobject_1;
    MoveL P1_3,v100,z1,MyNewTool\WObj:=Workobject_1;
    MoveL P1_4,v100,z1,MyNewTool\WObj:=Workobject_1;
    MoveL P1_5,v100,z1,MyNewTool\WObj:=Workobject_1;
    MoveL P1_6,v100,z1,MyNewTool\WObj:=Workobject_1;
    MoveL P1_7,v100,z1,MyNewTool\WObj:=Workobject_1;
    MoveL P1_8,v100,z1,MyNewTool\WObj:=Workobject_1;
    MoveL P1_9,v100,z1,MyNewTool\WObj:=Workobject_1;
    MoveL P1_10,v100,z1,MyNewTool\WObj:=Workobject_1;
    MoveL P1_11,v100,z1,MyNewTool\WObj:=Workobject_1;
    MoveL P1_12,v100,z1,MyNewTool\WObj:=Workobject_1;
    MoveL P1_13,v100,z1,MyNewTool\WObj:=Workobject_1;
    MoveL P1_14,v100,z1,MyNewTool\WObj:=Workobject_1;
    MoveL P1_15,v100,z1,MyNewTool\WObj:=Workobject_1;
    MoveL P1_16,v100,z1,MyNewTool\WObj:=Workobject_1;
    MoveL P1_17,v100,z1,MyNewTool\WObj:=Workobject_1;
    MoveL P1_18,v100,z1,MyNewTool\WObj:=Workobject_1;
    MoveL P1_19,v100,z1,MyNewTool\WObj:=Workobject_1;
    MoveL P1_20,v100,z1,MyNewTool\WObj:=Workobject_1;
    MoveL P1_21,v100,z1,MyNewTool\WObj:=Workobject_1;
    MoveL P1_22,v100,z1,MyNewTool\WObj:=Workobject_1;
    MoveL P1_23,v100,z1,MyNewTool\WObj:=Workobject_1;
    MoveL P1_24,v100,z1,MyNewTool\WObj:=Workobject_1;
    MoveL P1_25,v100,z1,MyNewTool\WObj:=Workobject_1;
    MoveL P1_26,v100,z1,MyNewTool\WObj:=Workobject_1;
    MoveL P1_27,v100,z1,MyNewTool\WObj:=Workobject_1;
    MoveL P1_28,v100,z1,MyNewTool\WObj:=Workobject_1;
    MoveL P1_29,v100,z1,MyNewTool\WObj:=Workobject_1;
    MoveL P1_30,v100,z1,MyNewTool\WObj:=Workobject_1;
    MoveL P1_31,v100,z1,MyNewTool\WObj:=Workobject_1;
    MoveL P1_32,v100,z1,MyNewTool\WObj:=Workobject_1;
    MoveL P1_33,v100,z1,MyNewTool\WObj:=Workobject_1;
    MoveL P1_34,v100,z1,MyNewTool\WObj:=Workobject_1;
    MoveL P1_35,v100,z1,MyNewTool\WObj:=Workobject_1;
    MoveL P1_36,v100,z1,MyNewTool\WObj:=Workobject_1;
    MoveL P1_37,v100,z1,MyNewTool\WObj:=Workobject_1;
    MoveL P1_38,v100,z1,MyNewTool\WObj:=Workobject_1;
    MoveL P1_39,v100,z1,MyNewTool\WObj:=Workobject_1;
    MoveL P1_40,v100,z1,MyNewTool\WObj:=Workobject_1;
    MoveL P1_41,v100,z1,MyNewTool\WObj:=Workobject_1;
    MoveL P1_42,v100,z1,MyNewTool\WObj:=Workobject_1;
    MoveL P1_43,v100,z1,MyNewTool\WObj:=Workobject_1;
    MoveL P1_44,v100,z1,MyNewTool\WObj:=Workobject_1;
    MoveL P1_45,v100,z1,MyNewTool\WObj:=Workobject_1;
    MoveL P1_46,v100,z1,MyNewTool\WObj:=Workobject_1;
    MoveL P1_47,v100,z1,MyNewTool\WObj:=Workobject_1;
    MoveL P1_48,v100,z1,MyNewTool\WObj:=Workobject_1;
    MoveL P1_49,v100,z1,MyNewTool\WObj:=Workobject_1;
    MoveL P1_50,v100,z1,MyNewTool\WObj:=Workobject_1;
    MoveL P1_51,v100,z1,MyNewTool\WObj:=Workobject_1;
    MoveL P1_52,v100,z1,MyNewTool\WObj:=Workobject_1;
    MoveL P1_53,v100,z1,MyNewTool\WObj:=Workobject_1;
    MoveL P1_54,v100,z1,MyNewTool\WObj:=Workobject_1;
    MoveL P1_55,v100,z1,MyNewTool\WObj:=Workobject_1;
    MoveL P1_56,v100,z1,MyNewTool\WObj:=Workobject_1;
    MoveL P1_57,v100,z1,MyNewTool\WObj:=Workobject_1;
    MoveL P1_58,v100,z1,MyNewTool\WObj:=Workobject_1;
    MoveL P1_59,v100,z1,MyNewTool\WObj:=Workobject_1;
    MoveL P1_60,v100,z1,MyNewTool\WObj:=Workobject_1;
    MoveL P1_61,v100,z1,MyNewTool\WObj:=Workobject_1;
    MoveL P1_62,v100,z1,MyNewTool\WObj:=Workobject_1;
    MoveL P1_63,v100,z1,MyNewTool\WObj:=Workobject_1;
    MoveL P1_64,v100,z1,MyNewTool\WObj:=Workobject_1;
    MoveL P1_65,v100,z1,MyNewTool\WObj:=Workobject_1;
    MoveL P1_66,v100,z1,MyNewTool\WObj:=Workobject_1;
    MoveL P1_67,v100,z1,MyNewTool\WObj:=Workobject_1;
    MoveL P1_68,v100,z1,MyNewTool\WObj:=Workobject_1;
    MoveL P1_69,v100,z1,MyNewTool\WObj:=Workobject_1;
    MoveL P1_70,v100,z1,MyNewTool\WObj:=Workobject_1;
    MoveL P1_71,v100,z1,MyNewTool\WObj:=Workobject_1;
    MoveL P1_72,v100,z1,MyNewTool\WObj:=Workobject_1;
    MoveL P1_73,v100,z1,MyNewTool\WObj:=Workobject_1;
    MoveL P1_74,v100,z1,MyNewTool\WObj:=Workobject_1;
    MoveL P1_75,v100,z1,MyNewTool\WObj:=Workobject_1;
    MoveL P1_76,v100,z1,MyNewTool\WObj:=Workobject_1;
    MoveL P1_77,v100,z1,MyNewTool\WObj:=Workobject_1;
    MoveL P1_78,v100,z1,MyNewTool\WObj:=Workobject_1;
    MoveL P1_79,v100,z1,MyNewTool\WObj:=Workobject_1;
    MoveL P1_80,v100,z1,MyNewTool\WObj:=Workobject_1;
    MoveL P1_81,v100,z1,MyNewTool\WObj:=Workobject_1;
    MoveL P1_82,v100,z1,MyNewTool\WObj:=Workobject_1;
    MoveL P1_83,v100,z1,MyNewTool\WObj:=Workobject_1;
    MoveL P1_84,v100,z1,MyNewTool\WObj:=Workobject_1;
    MoveL P1_85,v100,z1,MyNewTool\WObj:=Workobject_1;
    MoveL P1_86,v100,z1,MyNewTool\WObj:=Workobject_1;
    MoveL P1_87,v100,z1,MyNewTool\WObj:=Workobject_1;
    MoveL P1_88,v100,z1,MyNewTool\WObj:=Workobject_1;
    MoveL P1_89,v100,z1,MyNewTool\WObj:=Workobject_1;
    MoveL P1_90,v100,z1,MyNewTool\WObj:=Workobject_1;
    MoveL P1_91,v100,z1,MyNewTool\WObj:=Workobject_1;
    MoveL P1_92,v100,z1,MyNewTool\WObj:=Workobject_1;
    MoveL P1_93,v100,z1,MyNewTool\WObj:=Workobject_1;
    MoveL P1_94,v100,z1,MyNewTool\WObj:=Workobject_1;
    MoveL P1_95,v100,z1,MyNewTool\WObj:=Workobject_1;
    MoveL P1_96,v100,z1,MyNewTool\WObj:=Workobject_1;
    MoveL P1_97,v100,z1,MyNewTool\WObj:=Workobject_1;
    MoveL P1_98,v100,z1,MyNewTool\WObj:=Workobject_1;
    MoveL P1_99,v100,z1,MyNewTool\WObj:=Workobject_1;
    MoveL P1_100,v100,z1,MyNewTool\WObj:=Workobject_1;
    MoveL P1_101,v100,z1,MyNewTool\WObj:=Workobject_1;
    MoveL P1_102,v100,z1,MyNewTool\WObj:=Workobject_1;
    MoveL P1_103,v100,z1,MyNewTool\WObj:=Workobject_1;
    MoveL P1_104,v100,z1,MyNewTool\WObj:=Workobject_1;
    MoveL P1_105,v100,z1,MyNewTool\WObj:=Workobject_1;
    MoveL P1_106,v100,z1,MyNewTool\WObj:=Workobject_1;
    MoveL P1_107,v100,z1,MyNewTool\WObj:=Workobject_1;
    MoveL P1_108,v100,z1,MyNewTool\WObj:=Workobject_1;
    MoveL P1_109,v100,z1,MyNewTool\WObj:=Workobject_1;
    MoveL P1_110,v100,z1,MyNewTool\WObj:=Workobject_1;
    MoveL P1_111,v100,z1,MyNewTool\WObj:=Workobject_1;
    MoveL P1_112,v100,z1,MyNewTool\WObj:=Workobject_1;
    MoveL P1_113,v100,z1,MyNewTool\WObj:=Workobject_1;
    MoveL P1_114,v100,z1,MyNewTool\WObj:=Workobject_1;
    MoveL P1_115,v100,z1,MyNewTool\WObj:=Workobject_1;
    MoveL P1_116,v100,z1,MyNewTool\WObj:=Workobject_1;
    MoveL P1_117,v100,z1,MyNewTool\WObj:=Workobject_1;
    MoveL P1_118,v100,z1,MyNewTool\WObj:=Workobject_1;
    MoveL P1_119,v100,z1,MyNewTool\WObj:=Workobject_1;
    MoveL P1_120,v100,z1,MyNewTool\WObj:=Workobject_1;
    MoveL P1_121,v100,z1,MyNewTool\WObj:=Workobject_1;
    MoveL P1_122,v100,z1,MyNewTool\WObj:=Workobject_1;
    MoveL P1_123,v100,z1,MyNewTool\WObj:=Workobject_1;
    MoveL P1_124,v100,z1,MyNewTool\WObj:=Workobject_1;
    MoveL P1_125,v100,z1,MyNewTool\WObj:=Workobject_1;
    MoveL P1_126,v100,z1,MyNewTool\WObj:=Workobject_1;
    MoveL P1_127,v100,z1,MyNewTool\WObj:=Workobject_1;
    MoveL P1_128,v100,z1,MyNewTool\WObj:=Workobject_1;
    MoveL P1_129,v100,z1,MyNewTool\WObj:=Workobject_1;
    MoveL P1_130,v100,z1,MyNewTool\WObj:=Workobject_1;
    MoveL P1_131,v100,z1,MyNewTool\WObj:=Workobject_1;
    MoveL P1_132,v100,z1,MyNewTool\WObj:=Workobject_1;
    MoveL P1_133,v100,z1,MyNewTool\WObj:=Workobject_1;
    MoveL P1_134,v100,z1,MyNewTool\WObj:=Workobject_1;
    MoveL P1_135,v100,z1,MyNewTool\WObj:=Workobject_1;
    MoveL P1_136,v100,z1,MyNewTool\WObj:=Workobject_1;
    MoveL P1_137,v100,z1,MyNewTool\WObj:=Workobject_1;
    MoveL P1_138,v100,z1,MyNewTool\WObj:=Workobject_1;
    MoveL P1_139,v100,z1,MyNewTool\WObj:=Workobject_1;
    MoveL P1_140,v100,z1,MyNewTool\WObj:=Workobject_1;
    MoveL P1_141,v100,z1,MyNewTool\WObj:=Workobject_1;
    MoveL P1_142,v100,z1,MyNewTool\WObj:=Workobject_1;
    MoveL P1_143,v100,z1,MyNewTool\WObj:=Workobject_1;
    MoveL P1_144,v100,z1,MyNewTool\WObj:=Workobject_1;
    MoveL P1_145,v100,z1,MyNewTool\WObj:=Workobject_1;
    MoveL P1_146,v100,z1,MyNewTool\WObj:=Workobject_1;
    MoveL P1_147,v100,z1,MyNewTool\WObj:=Workobject_1;
    MoveL P1_148,v100,z1,MyNewTool\WObj:=Workobject_1;
    MoveL P1_149,v100,z1,MyNewTool\WObj:=Workobject_1;
    MoveL P1_150,v100,z1,MyNewTool\WObj:=Workobject_1;
    MoveL P1_151,v100,z1,MyNewTool\WObj:=Workobject_1;
    MoveL P1_152,v100,z1,MyNewTool\WObj:=Workobject_1;
    MoveL P1_153,v100,z1,MyNewTool\WObj:=Workobject_1;
    MoveL P1_154,v100,z1,MyNewTool\WObj:=Workobject_1;
    MoveL P1_1,v100,z1,MyNewTool\WObj:=Workobject_1;
    MoveL DibujoPk,v100,z1,MyNewTool\WObj:=Workobject_1;
  ENDPROC
  PROC Trazo2()
    MoveL DibujoPk,v100,z1,MyNewTool\WObj:=Workobject_1;
    MoveL P2_1,v100,z1,MyNewTool\WObj:=Workobject_1;
    MoveL P2_2,v100,z1,MyNewTool\WObj:=Workobject_1;
    MoveL P2_3,v100,z1,MyNewTool\WObj:=Workobject_1;
    MoveL P2_4,v100,z1,MyNewTool\WObj:=Workobject_1;
    MoveL P2_1,v100,z1,MyNewTool\WObj:=Workobject_1;
    MoveL DibujoPk,v100,z1,MyNewTool\WObj:=Workobject_1;
  ENDPROC
  PROC Trazo3()
    MoveL DibujoPk,v100,z1,MyNewTool\WObj:=Workobject_1;
    MoveL P3_1,v100,z1,MyNewTool\WObj:=Workobject_1;
    MoveL P3_2,v100,z1,MyNewTool\WObj:=Workobject_1;
    MoveL P3_3,v100,z1,MyNewTool\WObj:=Workobject_1;
    MoveL P3_4,v100,z1,MyNewTool\WObj:=Workobject_1;
    MoveL P3_5,v100,z1,MyNewTool\WObj:=Workobject_1;
    MoveL P3_6,v100,z1,MyNewTool\WObj:=Workobject_1;
    MoveL P3_7,v100,z1,MyNewTool\WObj:=Workobject_1;
    MoveL P3_8,v100,z1,MyNewTool\WObj:=Workobject_1;
    MoveL P3_1,v100,z1,MyNewTool\WObj:=Workobject_1;
    MoveL DibujoPk,v100,z1,MyNewTool\WObj:=Workobject_1;
  ENDPROC
  PROC Trazo4()
    MoveL DibujoPk,v100,z1,MyNewTool\WObj:=Workobject_1;
    MoveL P4_1,v100,z1,MyNewTool\WObj:=Workobject_1;
    MoveL P4_2,v100,z1,MyNewTool\WObj:=Workobject_1;
    MoveL P4_3,v100,z1,MyNewTool\WObj:=Workobject_1;
    MoveL P4_4,v100,z1,MyNewTool\WObj:=Workobject_1;
    MoveL P4_5,v100,z1,MyNewTool\WObj:=Workobject_1;
    MoveL P4_6,v100,z1,MyNewTool\WObj:=Workobject_1;
    MoveL P4_7,v100,z1,MyNewTool\WObj:=Workobject_1;
    MoveL P4_8,v100,z1,MyNewTool\WObj:=Workobject_1;
    MoveL P4_1,v100,z1,MyNewTool\WObj:=Workobject_1;
    MoveL DibujoPk,v100,z1,MyNewTool\WObj:=Workobject_1;
  ENDPROC
  PROC Trazo5()
    MoveL DibujoPk,v100,z1,MyNewTool\WObj:=Workobject_1;
    MoveL P5_1,v100,z1,MyNewTool\WObj:=Workobject_1;
    MoveL P5_2,v100,z1,MyNewTool\WObj:=Workobject_1;
    MoveL P5_3,v100,z1,MyNewTool\WObj:=Workobject_1;
    MoveL P5_4,v100,z1,MyNewTool\WObj:=Workobject_1;
    MoveL P5_1,v100,z1,MyNewTool\WObj:=Workobject_1;
    MoveL DibujoPk,v100,z1,MyNewTool\WObj:=Workobject_1;
  ENDPROC
  PROC Trazo6()
    MoveL DibujoPk,v100,z1,MyNewTool\WObj:=Workobject_1;
    MoveL P6_1,v100,z1,MyNewTool\WObj:=Workobject_1;
    MoveL P6_2,v100,z1,MyNewTool\WObj:=Workobject_1;
    MoveL P6_3,v100,z1,MyNewTool\WObj:=Workobject_1;
    MoveL P6_4,v100,z1,MyNewTool\WObj:=Workobject_1;
    MoveL P6_5,v100,z1,MyNewTool\WObj:=Workobject_1;
    MoveL P6_6,v100,z1,MyNewTool\WObj:=Workobject_1;
    MoveL P6_7,v100,z1,MyNewTool\WObj:=Workobject_1;
    MoveL P6_8,v100,z1,MyNewTool\WObj:=Workobject_1;
    MoveL P6_9,v100,z1,MyNewTool\WObj:=Workobject_1;
    MoveL P6_10,v100,z1,MyNewTool\WObj:=Workobject_1;
    MoveL P6_11,v100,z1,MyNewTool\WObj:=Workobject_1;
    MoveL P6_12,v100,z1,MyNewTool\WObj:=Workobject_1;
    MoveL P6_1,v100,z1,MyNewTool\WObj:=Workobject_1;
    MoveL DibujoPk,v100,z1,MyNewTool\WObj:=Workobject_1;
  ENDPROC
  PROC Trazo7()
    MoveL DibujoPk,v100,z1,MyNewTool\WObj:=Workobject_1;
    MoveL P7_1,v100,z1,MyNewTool\WObj:=Workobject_1;
    MoveL P7_2,v100,z1,MyNewTool\WObj:=Workobject_1;
    MoveL P7_3,v100,z1,MyNewTool\WObj:=Workobject_1;
    MoveL P7_4,v100,z1,MyNewTool\WObj:=Workobject_1;
    MoveL P7_5,v100,z1,MyNewTool\WObj:=Workobject_1;
    MoveL P7_6,v100,z1,MyNewTool\WObj:=Workobject_1;
    MoveL P7_7,v100,z1,MyNewTool\WObj:=Workobject_1;
    MoveL P7_8,v100,z1,MyNewTool\WObj:=Workobject_1;
    MoveL P7_9,v100,z1,MyNewTool\WObj:=Workobject_1;
    MoveL P7_10,v100,z1,MyNewTool\WObj:=Workobject_1;
    MoveL P7_11,v100,z1,MyNewTool\WObj:=Workobject_1;
    MoveL P7_12,v100,z1,MyNewTool\WObj:=Workobject_1;
    MoveL P7_1,v100,z1,MyNewTool\WObj:=Workobject_1;
    MoveL DibujoPk,v100,z1,MyNewTool\WObj:=Workobject_1;
  ENDPROC
  PROC Trazo8()
    MoveL DibujoPk,v100,z1,MyNewTool\WObj:=Workobject_1;
    MoveL P8_1,v100,z1,MyNewTool\WObj:=Workobject_1;
    MoveL P8_2,v100,z1,MyNewTool\WObj:=Workobject_1;
    MoveL P8_3,v100,z1,MyNewTool\WObj:=Workobject_1;
    MoveL P8_4,v100,z1,MyNewTool\WObj:=Workobject_1;
    MoveL P8_5,v100,z1,MyNewTool\WObj:=Workobject_1;
    MoveL P8_6,v100,z1,MyNewTool\WObj:=Workobject_1;
    MoveL P8_7,v100,z1,MyNewTool\WObj:=Workobject_1;
    MoveL P8_8,v100,z1,MyNewTool\WObj:=Workobject_1;
    MoveL P8_1,v100,z1,MyNewTool\WObj:=Workobject_1;
    MoveL DibujoPk,v100,z1,MyNewTool\WObj:=Workobject_1;
  ENDPROC
  PROC L()
    MoveJ L1,v100,z1,MyNewTool\WObj:=Workobject_1;
    MoveL L2,v100,z1,MyNewTool\WObj:=Workobject_1;
    MoveL L3,v100,z1,MyNewTool\WObj:=Workobject_1;
  ENDPROC
  PROC E_2()
    MoveJ E1_2,v100,z1,MyNewTool\WObj:=Workobject_1;
    MoveC E2_2,E3_2,v100,z1,MyNewTool\WObj:=Workobject_1;
    MoveC E4_2,E5_2,v100,z1,MyNewTool\WObj:=Workobject_1;
    MoveL E6_2,v100,z1,MyNewTool\WObj:=Workobject_1;
    MoveC E7_2,E5_2,v100,z1,MyNewTool\WObj:=Workobject_1;
  ENDPROC
  PROC O_2()
    MoveJ O1_2,v100,z1,MyNewTool\WObj:=Workobject_1;
    MoveC O2_2,O3_2,v100,z1,MyNewTool\WObj:=Workobject_1;
    MoveC O4_2,O1_2,v100,z1,MyNewTool\WObj:=Workobject_1;
  ENDPROC
  PROC N()
    MoveJ N1,v100,z1,MyNewTool\WObj:=Workobject_1;
    MoveL N2,v100,z1,MyNewTool\WObj:=Workobject_1;
    MoveC N3,N4,v100,z1,MyNewTool\WObj:=Workobject_1;
    MoveL N5,v100,z1,MyNewTool\WObj:=Workobject_1;
  ENDPROC
  PROC A()
    MoveJ A1,v100,z1,MyNewTool\WObj:=Workobject_1;
    MoveL A2,v100,z1,MyNewTool\WObj:=Workobject_1;
    MoveC A3,A4,v100,z1,MyNewTool\WObj:=Workobject_1;
    MoveJ Dibujo,v100,z1,MyNewTool\WObj:=Workobject_1;
    MoveJ A2,v100,z1,MyNewTool\WObj:=Workobject_1;
    MoveL A5,v100,z1,MyNewTool\WObj:=Workobject_1;
    MoveC A6,A7,v100,z1,MyNewTool\WObj:=Workobject_1;
    MoveC A8,A9,v100,z1,MyNewTool\WObj:=Workobject_1;
  ENDPROC
  PROC R()
    MoveJ R1,v100,z1,MyNewTool\WObj:=Workobject_1;
    MoveL R2,v100,z1,MyNewTool\WObj:=Workobject_1;
    MoveC R2_2,R3,v100,z1,MyNewTool\WObj:=Workobject_1;
  ENDPROC
  PROC D()
    MoveJ D1,v100,z1,MyNewTool\WObj:=Workobject_1;
    MoveC D2,D3,v100,z1,MyNewTool\WObj:=Workobject_1;
    MoveC D4,D1,v100,z1,MyNewTool\WObj:=Workobject_1;
    MoveJ Dibujo,v100,z1,MyNewTool\WObj:=Workobject_1;
    MoveJ D5,v100,z1,MyNewTool\WObj:=Workobject_1;
    MoveL D6,v100,z1,MyNewTool\WObj:=Workobject_1;
  ENDPROC
  PROC O_3()
    MoveJ O1_3,v100,z1,MyNewTool\WObj:=Workobject_1;
    MoveC O2_3,O3_3,v100,z1,MyNewTool\WObj:=Workobject_1;
    MoveC O4_3,O1_3,v100,z1,MyNewTool\WObj:=Workobject_1;
  ENDPROC
  PROC Home_F()
    MoveJ Dibujo,v100,z1,MyNewTool\WObj:=Workobject_1;
    MoveJ Home_2,v100,z1,MyNewTool\WObj:=Workobject_1;
    MoveJ Home,v100,z1,MyNewTool\WObj:=Workobject_1;
    MoveL RealH,v100,z1,MyNewTool\WObj:=Workobject_1;
  ENDPROC
  PROC Mantenimiento_p()
    MoveJ Home_F2,v100,z1,MyNewTool\WObj:=Workobject_1;
    MoveJ Mantenimiento,v100,z1,MyNewTool\WObj:=Workobject_1;
  ENDPROC
  PROC Home_F_2()
    MoveJ Home_F2,v100,z1,MyNewTool\WObj:=Workobject_1;
  ENDPROC
  PROC Home_0()
    MoveJ Home0,v100,z1,MyNewTool\WObj:=Workobject_1;
  ENDPROC
  PROC Aura()
    MoveJ Aura0,v200,z1,MyNewTool\WObj:=Workobject_1;
    MoveJ Aura1,v200,z1,MyNewTool\WObj:=Workobject_1;
    MoveJ Aura2,v200,z1,MyNewTool\WObj:=Workobject_1;
    MoveJ Aura3,v200,z1,MyNewTool\WObj:=Workobject_1;
    MoveJ Aura4,v200,z1,MyNewTool\WObj:=Workobject_1;
    MoveJ Aura5,v200,z1,MyNewTool\WObj:=Workobject_1;
    MoveJ Aura6,v200,z1,MyNewTool\WObj:=Workobject_1;
    MoveJ Aura7,v200,z1,MyNewTool\WObj:=Workobject_1;
    MoveJ Aura8,v200,z1,MyNewTool\WObj:=Workobject_1;
    MoveJ Aura1,v200,z1,MyNewTool\WObj:=Workobject_1;
  ENDPROC
  PROC Real_Home()
    MoveJ RealH,v100,z1,MyNewTool\WObj:=Workobject_1;
  ENDPROC
  PROC Posicionar_Banda()
    Reset FWD_Conveyor;
    Reset BWD_Conveyor;
    Set BWD_Conveyor;
    WaitTime 2.591;
    Reset BWD_Conveyor;
  ENDPROC
ENDMODULE

! task T_ROB1
MODULE Pikachu
  LOCAL CONST robtarget OrigenPikachu:=[[73.025,-352.375,-150],[0,0.707106781,0.707106781,0],[0,0,0,0],[9E+09,9E+09,9E+09,9E+09,9E+09,9E+09]];
ENDMODULE

